{attribute 'Tc2GvlVarNames'}
VAR_GLOBAL
		tPLC_TaskCycleTime_ms			:TIME 	:=	LREAL_TO_TIME(GVL.lrgActCycleTime * 1000) ;		(* PLC Task Cycle Time in [ms] *)
END_VAR

(* stored: Version 1.1.0.1, ProductVersion 3.1.4024.15
   GVL GVL_Gr00Init: Id {db7b2612-5963-46a8-9be5-b4c0dded8796} *)
